// TIA Portal V20 export
// export: Created 2026-10-20T12:56:13.3503517Z, ExportSetting WithDefaults, DisplayName Totally Integrated Automation Portal, DisplayVersion V20 Update 6, DisplayName TIA Portal Openness, DisplayVersion V20 Update 6, DisplayName TIA Portal Version Control Interface, DisplayVersion V20 Update 6, DisplayName SINAMICS Startdrive Advanced, DisplayVersion V20 SP1, DisplayName SINAMICS Startdrive G130, G150, S120, S150, SINAMICS MV, G220, S200, S210, DisplayVersion V20 SP1, DisplayName SINAMICS Startdrive G110M, G120, G120C, G120D, G120P, G115D, DisplayVersion V20 SP1, DisplayName STEP 7 Professional, DisplayVersion V20 Update 6, DisplayName STEP 7 Safety, DisplayVersion V20 Update 2, DisplayName WinCC Basic/Comfort/Advanced, DisplayVersion V20 Update 6, DisplayName WinCC Unified, DisplayVersion V20 Update 6
DATA_BLOCK "Shuttle_TCP_Comms_FB_DB_1"   // DB64
VERSION : 0.1
// stored: AutoNumber true, DBAccessibleFromOPCUA true, InstanceOfName Shuttle_TCP_Comms, InstanceOfType FB
"Shuttle_TCP_Comms"
   // VAR_INPUT
   //    Enable : Bool;
   //    "E-stop" : Bool;
   //    TCP_Configuration : "LCom_typeConfig";
   //    Shuttle_No : UInt;
   // END_VAR
   // VAR_OUTPUT
   //    Connected : Bool;
   //    Busy : Bool;
   //    Status : Word;
   //    Error : Bool;
   // END_VAR
   // VAR_IN_OUT
   //    TCP_Diag : "LCom_typeDiagnostics";
   //    LCom_Communication_DB : "LCom_Communication_FB";
   // END_VAR
   // VAR
   //    SendBuffer { ExternalAccessible := 'False'; ExternalVisible := 'False'; ExternalWritable := 'False'} : Array[0..6] of Byte;
   //    ReceiveBuffer { ExternalAccessible := 'False'; ExternalVisible := 'False'; ExternalWritable := 'False'} : Array[0..1] of Byte;
   //    Send : Bool;
   //    SendDataLength : USInt;
   //    Sending : Bool;
   //    T_Send_DB { S7_SetPoint := 'True'} : TON_TIME;
   // END_VAR
BEGIN
END_DATA_BLOCK
